FUNCTION_BLOCK CONVEYOR_INTERLOCK (* Migrated from IEC 61131-3 ST *)
  (* Standard: 61499-2 *)
  (* Version 1.0, 2026-11-06, st2fb *)
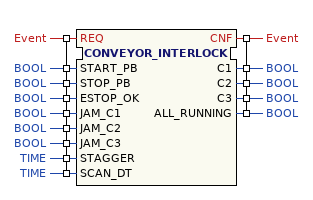
  EVENT_INPUT
    REQ WITH START_PB, STOP_PB, ESTOP_OK, JAM_C1, JAM_C2, JAM_C3, STAGGER, SCAN_DT;
  END_EVENT
  EVENT_OUTPUT
    CNF WITH C1, C2, C3, ALL_RUNNING;
  END_EVENT
  VAR_INPUT
    START_PB : BOOL;
    STOP_PB : BOOL;
    ESTOP_OK : BOOL;
    JAM_C1 : BOOL;
    JAM_C2 : BOOL;
    JAM_C3 : BOOL;
    STAGGER : TIME;
    SCAN_DT : TIME;
  END_VAR
  VAR_OUTPUT
    C1 : BOOL;
    C2 : BOOL;
    C3 : BOOL;
    ALL_RUNNING : BOOL;
  END_VAR
  VAR
    RUN_REQ : BOOL := FALSE;
    C1_CMD : BOOL := FALSE;
    C2_CMD : BOOL := FALSE;
    ST2FB_NOW : TIME := T#0s;
    ON_C2_IN : BOOL := FALSE;
    ON_C2_PT : TIME := T#0s;
    ON_C2_Q : BOOL := FALSE;
    ON_C2_ET : TIME := T#0s;
    ON_C2_STATE : INT := 0;
    ON_C2_PREV_IN : BOOL := FALSE;
    ON_C2_START_TIME : TIME := T#0s;
    ON_C1_IN : BOOL := FALSE;
    ON_C1_PT : TIME := T#0s;
    ON_C1_Q : BOOL := FALSE;
    ON_C1_ET : TIME := T#0s;
    ON_C1_STATE : INT := 0;
    ON_C1_PREV_IN : BOOL := FALSE;
    ON_C1_START_TIME : TIME := T#0s;
    CLEAR_C2_IN : BOOL := FALSE;
    CLEAR_C2_PT : TIME := T#0s;
    CLEAR_C2_Q : BOOL := FALSE;
    CLEAR_C2_ET : TIME := T#0s;
    CLEAR_C2_STATE : INT := 0;
    CLEAR_C2_PREV_IN : BOOL := FALSE;
    CLEAR_C2_START_TIME : TIME := T#0s;
    CLEAR_C3_IN : BOOL := FALSE;
    CLEAR_C3_PT : TIME := T#0s;
    CLEAR_C3_Q : BOOL := FALSE;
    CLEAR_C3_ET : TIME := T#0s;
    CLEAR_C3_STATE : INT := 0;
    CLEAR_C3_PREV_IN : BOOL := FALSE;
    CLEAR_C3_START_TIME : TIME := T#0s;
  END_VAR
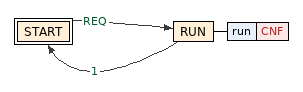
  EC_STATES
    START;
    RUN : run -> CNF;
  END_STATES
  EC_TRANSITIONS
    START TO RUN := REQ;
    RUN TO START := 1;
  END_TRANSITIONS
  ALGORITHM run IN ST:
ST2FB_NOW := ST2FB_NOW + SCAN_DT;
IF STOP_PB OR NOT ESTOP_OK OR JAM_C1 OR JAM_C2 OR JAM_C3 THEN
  RUN_REQ := FALSE;
ELSIF START_PB THEN
  RUN_REQ := TRUE;
END_IF;

ON_C2_IN := RUN_REQ;
ON_C2_PT := STAGGER;
IF (ON_C2_STATE = 0) AND NOT ON_C2_PREV_IN AND ON_C2_IN THEN
  ON_C2_STATE := 1;
  ON_C2_Q := FALSE;
  ON_C2_START_TIME := ST2FB_NOW;
ELSE
  IF NOT ON_C2_IN THEN
    ON_C2_ET := T#0s;
    ON_C2_Q := FALSE;
    ON_C2_STATE := 0;
  ELSIF ON_C2_STATE = 1 THEN
    IF ON_C2_START_TIME + ON_C2_PT <= ST2FB_NOW THEN
      ON_C2_STATE := 2;
      ON_C2_Q := TRUE;
      ON_C2_ET := ON_C2_PT;
    ELSE
      ON_C2_ET := ST2FB_NOW - ON_C2_START_TIME;
    END_IF;
  END_IF;
END_IF;
ON_C2_PREV_IN := ON_C2_IN;

ON_C1_IN := ON_C2_Q;
ON_C1_PT := STAGGER;
IF (ON_C1_STATE = 0) AND NOT ON_C1_PREV_IN AND ON_C1_IN THEN
  ON_C1_STATE := 1;
  ON_C1_Q := FALSE;
  ON_C1_START_TIME := ST2FB_NOW;
ELSE
  IF NOT ON_C1_IN THEN
    ON_C1_ET := T#0s;
    ON_C1_Q := FALSE;
    ON_C1_STATE := 0;
  ELSIF ON_C1_STATE = 1 THEN
    IF ON_C1_START_TIME + ON_C1_PT <= ST2FB_NOW THEN
      ON_C1_STATE := 2;
      ON_C1_Q := TRUE;
      ON_C1_ET := ON_C1_PT;
    ELSE
      ON_C1_ET := ST2FB_NOW - ON_C1_START_TIME;
    END_IF;
  END_IF;
END_IF;
ON_C1_PREV_IN := ON_C1_IN;

C1_CMD := ON_C1_Q;

CLEAR_C2_IN := C1_CMD;
CLEAR_C2_PT := STAGGER;
IF (CLEAR_C2_STATE = 0) AND CLEAR_C2_PREV_IN AND NOT CLEAR_C2_IN THEN
  CLEAR_C2_STATE := 1;
  CLEAR_C2_START_TIME := ST2FB_NOW;
ELSE
  IF CLEAR_C2_IN THEN
    CLEAR_C2_ET := T#0s;
    CLEAR_C2_STATE := 0;
  ELSIF CLEAR_C2_STATE = 1 THEN
    IF CLEAR_C2_START_TIME + CLEAR_C2_PT <= ST2FB_NOW THEN
      CLEAR_C2_STATE := 2;
      CLEAR_C2_ET := CLEAR_C2_PT;
    ELSE
      CLEAR_C2_ET := ST2FB_NOW - CLEAR_C2_START_TIME;
    END_IF;
  END_IF;
END_IF;
CLEAR_C2_Q := CLEAR_C2_IN OR (CLEAR_C2_STATE = 1);
CLEAR_C2_PREV_IN := CLEAR_C2_IN;

C2_CMD := ON_C2_Q OR CLEAR_C2_Q;

CLEAR_C3_IN := C2_CMD;
CLEAR_C3_PT := STAGGER;
IF (CLEAR_C3_STATE = 0) AND CLEAR_C3_PREV_IN AND NOT CLEAR_C3_IN THEN
  CLEAR_C3_STATE := 1;
  CLEAR_C3_START_TIME := ST2FB_NOW;
ELSE
  IF CLEAR_C3_IN THEN
    CLEAR_C3_ET := T#0s;
    CLEAR_C3_STATE := 0;
  ELSIF CLEAR_C3_STATE = 1 THEN
    IF CLEAR_C3_START_TIME + CLEAR_C3_PT <= ST2FB_NOW THEN
      CLEAR_C3_STATE := 2;
      CLEAR_C3_ET := CLEAR_C3_PT;
    ELSE
      CLEAR_C3_ET := ST2FB_NOW - CLEAR_C3_START_TIME;
    END_IF;
  END_IF;
END_IF;
CLEAR_C3_Q := CLEAR_C3_IN OR (CLEAR_C3_STATE = 1);
CLEAR_C3_PREV_IN := CLEAR_C3_IN;

C1 := C1_CMD AND ESTOP_OK AND NOT JAM_C1 AND NOT JAM_C2 AND NOT JAM_C3;
C2 := C2_CMD AND ESTOP_OK AND NOT JAM_C2 AND NOT JAM_C3;
C3 := (RUN_REQ OR CLEAR_C3_Q) AND ESTOP_OK AND NOT JAM_C3;
ALL_RUNNING := C1 AND C2 AND C3;
  END_ALGORITHM
END_FUNCTION_BLOCK
